(* IEC 61131-3 sources: ia2/examples/retain_recovery/pous, 1 file *)

(* ---- main.st ---- *)
PROGRAM main
VAR RETAIN value : DINT := 42; END_VAR
END_PROGRAM
